// TIA Portal V18 export
ORGANIZATION_BLOCK "OB1 Main"   // OB1, LAD, ProgramCycle
TITLE = "Main Program Sweep (Cycle)"
{ S7_Optimized_Access := 'TRUE' }
// stored: SetENOAutomatically false
   VAR_INPUT
      Initial_Call : Bool;   // Initial call of this OB
      Remanence : Bool;   // =True, if remanent data are available
   END_VAR
   VAR_TEMP
      ADR : UDInt;
      LEN : UInt;
      "RETURN" : Int;
      ERROR : Bool;
      STATUS : Word;
      DONE : Bool;
      POPID : String;
      CU : Int;
      Quantidade_erro : Int;
      DONE_MAIN_LINE_PUT : Bool;
      ERROR_MAIN_LINE_PUT : Bool;
      DONE_MAIN_LINE_GET : Bool;
      ERROR_MAIN_LINE_GET : Bool;
      DONE_FALCARE_PUT : Bool;
      ERROR_FALCARE_PUT : Bool;
      DONE_FALCARE_GET : Bool;
      ERROR_FALCARE_GET : Bool;
      DONE_GIRADOR_PUT : Bool;
      ERROR_GIRADOR_PUT : Bool;
      DONE_GIRADOR_GET : Bool;
      ERROR_GIRADOR_GET : Bool;
      DONE_ABSTECIMENTO_OLEO_PUT : Bool;
      ERRO_ABASTECIMENTO_OLEO_PUT : Bool;
      DONE_ABSTECIMENTO_OLEO_GET : Bool;
      ERRO_ABSTECIMENTO_OLEO_GET : Bool;
      ERROR_ALARMS_IHM_FALCARE_GET : Bool;
      DONE_ALARMS_IHM_FALCARE_GET : Bool;
      AUX_BSEND_LEMARB : Word;
      AUX_RECIVE_LEMARB : Word;
   END_VAR
BEGIN

REGION Network 1: Set Id Connection automatic
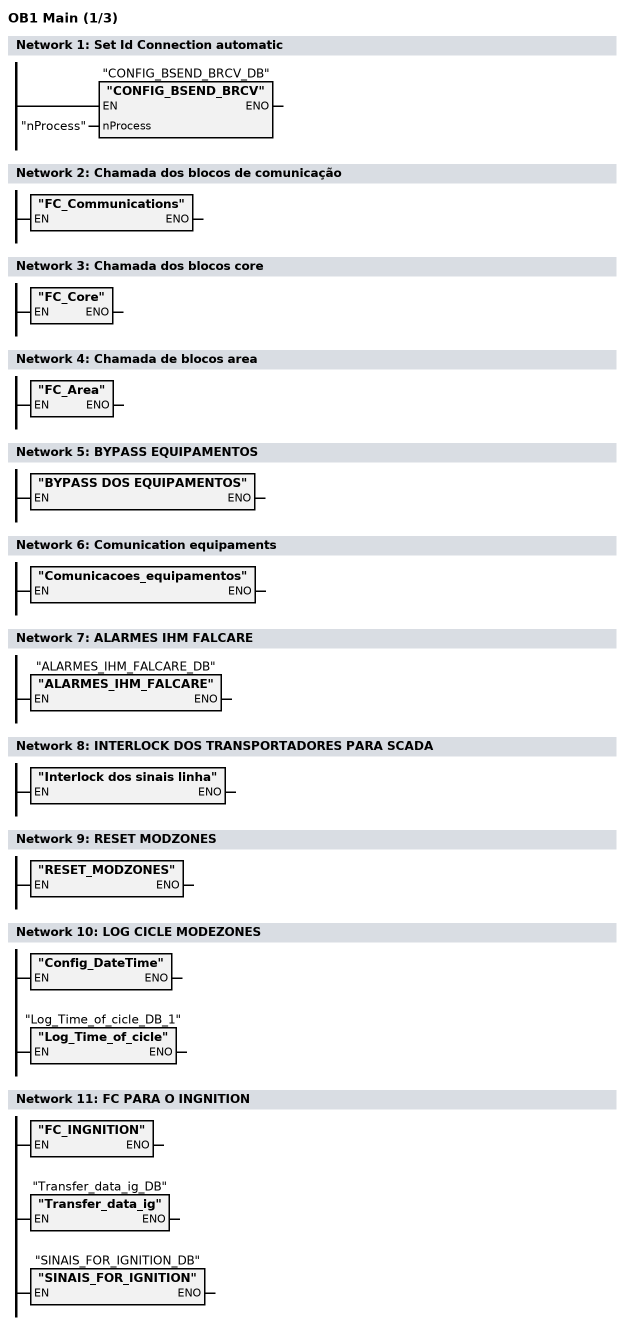
   RUNG wire#powerrail
      "CONFIG_BSEND_BRCV_DB"(nProcess := "nProcess")
   END_RUNG
   // the same network as SCL:
   "CONFIG_BSEND_BRCV_DB"(nProcess := "nProcess");   // "CONFIG_BSEND_BRCV"
END_REGION

REGION Network 2: Chamada dos blocos de comunicação
   RUNG wire#powerrail
      "FC_Communications"()
   END_RUNG
   // the same network as SCL:
   "FC_Communications"();
END_REGION

REGION Network 3: Chamada dos blocos core
   RUNG wire#powerrail
      "FC_Core"()
   END_RUNG
   // the same network as SCL:
   "FC_Core"();
END_REGION

REGION Network 4: Chamada de blocos area
   RUNG wire#powerrail
      "FC_Area"()
   END_RUNG
   // the same network as SCL:
   "FC_Area"();
END_REGION

REGION Network 5: BYPASS EQUIPAMENTOS
   RUNG wire#powerrail
      "BYPASS DOS EQUIPAMENTOS"()
   END_RUNG
   // the same network as SCL:
   "BYPASS DOS EQUIPAMENTOS"();
END_REGION

REGION Network 6: Comunication equipaments
   RUNG wire#powerrail
      "Comunicacoes_equipamentos"()
   END_RUNG
   // the same network as SCL:
   "Comunicacoes_equipamentos"();
END_REGION

REGION Network 7: ALARMES IHM FALCARE
   RUNG wire#powerrail
      "ALARMES_IHM_FALCARE_DB"()
   END_RUNG
   // the same network as SCL:
   "ALARMES_IHM_FALCARE_DB"();   // "ALARMES_IHM_FALCARE"
END_REGION

REGION Network 8: INTERLOCK DOS TRANSPORTADORES PARA SCADA
   RUNG wire#powerrail
      "Interlock dos sinais linha"()
   END_RUNG
   // the same network as SCL:
   "Interlock dos sinais linha"();
END_REGION

REGION Network 9: RESET MODZONES
   RUNG wire#powerrail
      "RESET_MODZONES"()
   END_RUNG
   // the same network as SCL:
   "RESET_MODZONES"();
END_REGION

REGION Network 10: LOG CICLE MODEZONES
   RUNG wire#powerrail
      "Config_DateTime"()
   END_RUNG
   RUNG wire#powerrail
      "Log_Time_of_cicle_DB_1"()
   END_RUNG
   // the same network as SCL:
   "Config_DateTime"();
   "Log_Time_of_cicle_DB_1"();   // "Log_Time_of_cicle"
END_REGION

REGION Network 11: FC PARA O INGNITION
   RUNG wire#powerrail
      "FC_INGNITION"()
   END_RUNG
   RUNG wire#powerrail
      "Transfer_data_ig_DB"()
   END_RUNG
   RUNG wire#powerrail
      "SINAIS_FOR_IGNITION_DB"()
   END_RUNG
   // the same network as SCL:
   "FC_INGNITION"();
   "Transfer_data_ig_DB"();   // "Transfer_data_ig"
   "SINAIS_FOR_IGNITION_DB"();   // "SINAIS_FOR_IGNITION"
END_REGION

REGION Network 12: TESTE DE VALIDAÇÃO MODEZONES
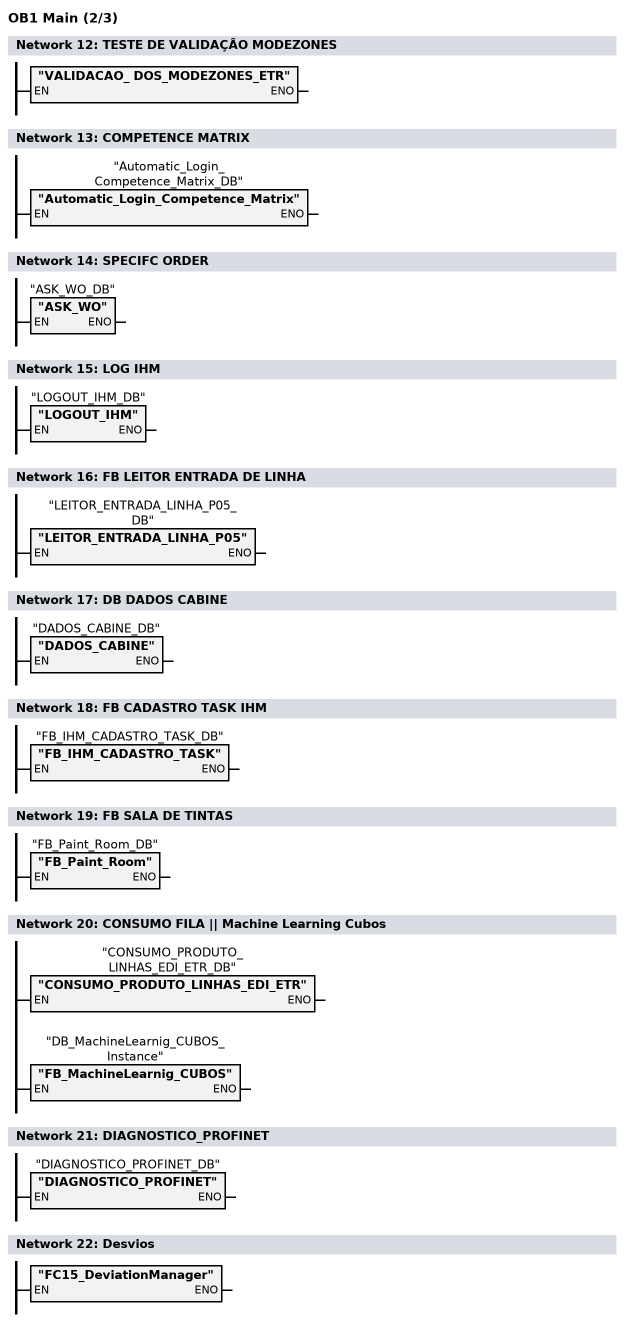
   RUNG wire#powerrail
      "VALIDACAO_ DOS_MODEZONES_ETR"()
   END_RUNG
   // the same network as SCL:
   "VALIDACAO_ DOS_MODEZONES_ETR"();
END_REGION

REGION Network 13: COMPETENCE MATRIX
   RUNG wire#powerrail
      "Automatic_Login_Competence_Matrix_DB"()
   END_RUNG
   // the same network as SCL:
   "Automatic_Login_Competence_Matrix_DB"();   // "Automatic_Login_Competence_Matrix"
END_REGION

REGION Network 14: SPECIFC ORDER
   RUNG wire#powerrail
      "ASK_WO_DB"()
   END_RUNG
   // the same network as SCL:
   "ASK_WO_DB"();   // "ASK_WO"
END_REGION

REGION Network 15: LOG IHM
   RUNG wire#powerrail
      "LOGOUT_IHM_DB"()
   END_RUNG
   // the same network as SCL:
   "LOGOUT_IHM_DB"();   // "LOGOUT_IHM"
END_REGION

REGION Network 16: FB LEITOR ENTRADA DE LINHA
   RUNG wire#powerrail
      "LEITOR_ENTRADA_LINHA_P05_DB"()
   END_RUNG
   // the same network as SCL:
   "LEITOR_ENTRADA_LINHA_P05_DB"();   // "LEITOR_ENTRADA_LINHA_P05"
END_REGION

REGION Network 17: DB DADOS CABINE
   RUNG wire#powerrail
      "DADOS_CABINE_DB"()
   END_RUNG
   // the same network as SCL:
   "DADOS_CABINE_DB"();   // "DADOS_CABINE"
END_REGION

REGION Network 18: FB CADASTRO TASK IHM
   RUNG wire#powerrail
      "FB_IHM_CADASTRO_TASK_DB"()
   END_RUNG
   // the same network as SCL:
   "FB_IHM_CADASTRO_TASK_DB"();   // "FB_IHM_CADASTRO_TASK"
END_REGION

REGION Network 19: FB SALA DE TINTAS
   RUNG wire#powerrail
      "FB_Paint_Room_DB"()
   END_RUNG
   // the same network as SCL:
   "FB_Paint_Room_DB"();   // "FB_Paint_Room"
END_REGION

REGION Network 20: CONSUMO FILA || Machine Learning Cubos
   RUNG wire#powerrail
      "CONSUMO_PRODUTO_LINHAS_EDI_ETR_DB"()
   END_RUNG
   RUNG wire#powerrail
      "DB_MachineLearnig_CUBOS_Instance"()
   END_RUNG
   // the same network as SCL:
   "CONSUMO_PRODUTO_LINHAS_EDI_ETR_DB"();   // "CONSUMO_PRODUTO_LINHAS_EDI_ETR"
   "DB_MachineLearnig_CUBOS_Instance"();   // "FB_MachineLearnig_CUBOS"
END_REGION

REGION Network 21: DIAGNOSTICO_PROFINET
   RUNG wire#powerrail
      "DIAGNOSTICO_PROFINET_DB"()
   END_RUNG
   // the same network as SCL:
   "DIAGNOSTICO_PROFINET_DB"();   // "DIAGNOSTICO_PROFINET"
END_REGION

REGION Network 22: Desvios
   RUNG wire#powerrail
      "FC15_DeviationManager"()
   END_RUNG
   // the same network as SCL:
   "FC15_DeviationManager"();
END_REGION

REGION Network 23: BSEND SEQUENCE NOW MD1
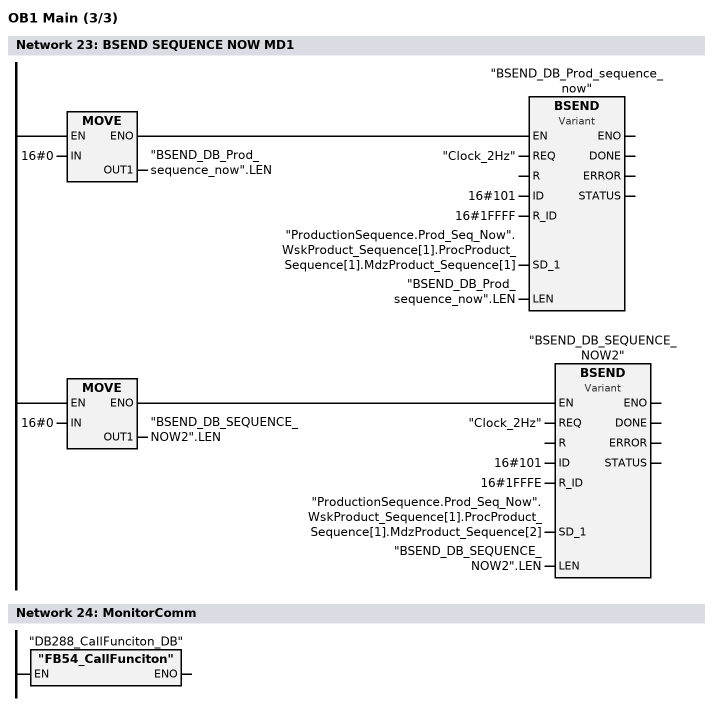
   RUNG wire#powerrail
      Move(in := 16#0, out1 => "BSEND_DB_Prod_sequence_now".LEN)
      { S7_Templates := "[ptr_type := Variant, id_type := CONN_PRG, r_id_type := CONN_R_ID]" } "BSEND_DB_Prod_sequence_now".BSEND(REQ := "Clock_2Hz", R :=, ID := 16#101, R_ID := 16#1FFFF, SD_1 := "ProductionSequence.Prod_Seq_Now".WskProduct_Sequence[1].ProcProduct_Sequence[1].MdzProduct_Sequence[1], LEN := "BSEND_DB_Prod_sequence_now".LEN, DONE =>, ERROR =>, STATUS =>)
   END_RUNG
   RUNG wire#powerrail
      Move(in := 16#0, out1 => "BSEND_DB_SEQUENCE_NOW2".LEN)
      { S7_Templates := "[ptr_type := Variant, id_type := CONN_PRG, r_id_type := CONN_R_ID]" } "BSEND_DB_SEQUENCE_NOW2".BSEND(REQ := "Clock_2Hz", R :=, ID := 16#101, R_ID := 16#1FFFE, SD_1 := "ProductionSequence.Prod_Seq_Now".WskProduct_Sequence[1].ProcProduct_Sequence[1].MdzProduct_Sequence[2], LEN := "BSEND_DB_SEQUENCE_NOW2".LEN, DONE =>, ERROR =>, STATUS =>)
   END_RUNG
   // the same network as SCL:
   "BSEND_DB_Prod_sequence_now".LEN := 16#0;
   "BSEND_DB_Prod_sequence_now"(REQ := "Clock_2Hz",   // BSEND
                           ID := 16#101,
                           R_ID := 16#1FFFF,
                           SD_1 := "ProductionSequence.Prod_Seq_Now".WskProduct_Sequence[1].ProcProduct_Sequence[1].MdzProduct_Sequence[1],
                           LEN := "BSEND_DB_Prod_sequence_now".LEN);
   "BSEND_DB_SEQUENCE_NOW2".LEN := 16#0;
   "BSEND_DB_SEQUENCE_NOW2"(REQ := "Clock_2Hz",   // BSEND
                           ID := 16#101,
                           R_ID := 16#1FFFE,
                           SD_1 := "ProductionSequence.Prod_Seq_Now".WskProduct_Sequence[1].ProcProduct_Sequence[1].MdzProduct_Sequence[2],
                           LEN := "BSEND_DB_SEQUENCE_NOW2".LEN);
END_REGION

REGION Network 24: MonitorComm
   RUNG wire#powerrail
      "DB288_CallFunciton_DB"()
   END_RUNG
   // the same network as SCL:
   "DB288_CallFunciton_DB"();   // "FB54_CallFunciton"
END_REGION
END_ORGANIZATION_BLOCK
